Fanuc KAREL source: KT00488.KL

PROGRAM KT00488
%NOLOCKGROUP
VAR
  P1: POSITION
  P2: JOINTPOS
  OUT: BOOLEAN
BEGIN
  OUT = P1 >=< P2
END KT00488
